Fanuc KAREL source: kt00327.KL

PROGRAM KT00327
%STACKSIZE=65535
%PRIORITY=65535
%NOLOCKGROUP
VAR
V1 : VECTOR
V2 : VECTOR
OUT : BOOLEAN
BEGIN
V1.X=1.0
V2.Y=2.0
V1.X=1.0
V2.Y=2.0
-- UNRESOLVED_PC line 12 opcodes [49 49 96 23] marker_code=80
END KT00327
